// TIA Portal V20 export
// export: Created 2026-10-19T18:02:47.4030367Z, ExportSetting WithDefaults, DisplayName Totally Integrated Automation Portal, DisplayVersion V20 Update 6, DisplayName TIA Portal Openness, DisplayVersion V20 Update 6, DisplayName TIA Portal Version Control Interface, DisplayVersion V20 Update 6, DisplayName SINAMICS Startdrive Advanced, DisplayVersion V20 SP1, DisplayName SINAMICS Startdrive G130, G150, S120, S150, SINAMICS MV, G220, S200, S210, DisplayVersion V20 SP1, DisplayName SINAMICS Startdrive G110M, G120, G120C, G120D, G120P, G115D, DisplayVersion V20 SP1, DisplayName STEP 7 Professional, DisplayVersion V20 Update 6, DisplayName STEP 7 Safety, DisplayVersion V20 Update 2, DisplayName WinCC Basic/Comfort/Advanced, DisplayVersion V20 Update 6, DisplayName WinCC Unified, DisplayVersion V20 Update 6
DATA_BLOCK "Control_DB"   // DB69
{ S7_Optimized_Access := 'TRUE' }
VERSION : 0.1
// stored: AutoNumber true, DBAccessibleFromOPCUA true, DBAccessibleFromWebserver true, IsOnlyStoredInLoadMemory false, IsRetainMemResEnabled false, IsWriteProtectedInAS false, MemoryReserve 100
   VAR
      Inbound_Cnv : "Inbound_Cnv_Control_UDT";
      PopUp_Cnv { S7_SetPoint := 'True'} : Array[1..4] of "PopUp_Cnv_Control";
      Outbound_Cnv { S7_SetPoint := 'True'} : "Outbound_Cnv_Control";
      ECnv_Control { S7_SetPoint := 'True'} : "ECnv_Control";
      LCnv_Control { S7_SetPoint := 'True'} : Array[1..3] of "Buffer_Cnv_Control";
      VTD_Control { S7_SetPoint := 'True'} : "VTD_Control";
      "VTD_Order Table" { S7_SetPoint := 'True'} : "WMS_OPC_UA";
      "Carrousel_Order Table" { S7_SetPoint := 'True'} : "WMS_OPC_UA";
      Shuttles_Position : Array[1..3] of Struct
         x : DInt;
         y : DInt;
         Charging : Bool;
      END_STRUCT;
      "Weighing Station" : Struct
         Start : Bool;
         Ready : Bool;
         Running : Bool;
         Done : Bool;
         Valid : Bool;
         Weight : Real;
         Error_ID : Word;
      END_STRUCT;
      "Profiling Station" : Struct
         Start : Bool;
         Ready : Bool;
         Running : Bool;
         Done : Bool;
         Valid : Bool;
         OverWidth : Bool;
         OverHeight : Bool;
         OverLength : Bool;
         Error_ID : Word;
      END_STRUCT;
      Pick_Station : Struct
         Cnv_Occupied { ExternalWritable := 'False'} : Bool;
         PushButton : Bool;
         LightGuard : Bool;
         PushButtonLight : Bool;
         Mode { ExternalWritable := 'False'} : UInt;
         Error { ExternalWritable := 'False'} : Bool;
         Warning { ExternalWritable := 'False'} : UInt;
         Enabled { ExternalWritable := 'False'} : Bool;
         Stopped { ExternalWritable := 'False'} : Bool;
         Done : Bool;
         Running { ExternalWritable := 'False'} : Bool;
         Ready_For_Task { ExternalWritable := 'False'} : Bool;
         Current_Task_Type : UInt;
         Current_Task_ID { ExternalWritable := 'False'} : UInt;
         Pallet_Type { ExternalWritable := 'False'} : UInt;
         SM_State { ExternalWritable := 'False'} : UInt;
         Motor : "Cnv_Motor";
         Instruction : "OutCnv_Instruction";
         Cnv_Errors { S7_SetPoint := 'True'} : "Cnv_Errors";
      END_STRUCT;
      InBarcode_Station : Struct
         Start : Bool;
         Ready : Bool;
         Running : Bool;
         Done : Bool;
         Valid : Bool;
         Barcode : String;
         "Reading Gate number" : String;
         "Reading Gate number OLD" : String;
         "Number of Reading Gates" : String;
         "Number of Reading Gates OLD" : String;
      END_STRUCT;
      OutBarcode_Station : Struct
         Start : Bool;
         Ready : Bool;
         Running : Bool;
         Done : Bool;
         Valid : Bool;
         Barcode : String;
         Barcode_Old : Array[1..16] of Char;
      END_STRUCT;
      VTDBarcode_Station : Struct
         Start : Bool;
         Ready : Bool;
         Running : Bool;
         Done : Bool;
         Valid : Bool;
         Barcode : String;
         Barcode_Old : String;
      END_STRUCT;
      Movement_Completed : Struct
         RTR_ITP1 : Bool;
         RTR_P1TP2 : Bool;
         RTR_P2TP3 : Bool;
         RTR_P3TP4 : Bool;
         RTR_P4TO : Bool;
         Chain_To_Chain : Bool;
         Pop4_To_Pick : Bool;
         Pick_To_Pop1 : Bool;
         WeighingStation : Bool;
      END_STRUCT;
   END_VAR
BEGIN
END_DATA_BLOCK
